(* IEC 61131-3 sources: codesys-framework/txt/application/WeVe Core (library)/30 Module/FB_Module/Properties, 4 files *)

(* ---- Busy.prop.st ---- *)
PROPERTY Busy : BOOL

// --- BEGIN IMPLEMENTATION ---

// ----------- GET -----------
VAR
END_VAR

// -- BEGIN IMPLEMENTATION GET --
Busy := _xBusy;

(* ---- Enabled.prop.st ---- *)
PROPERTY Enabled : BOOL

// --- BEGIN IMPLEMENTATION ---

// ----------- GET -----------
VAR
END_VAR

// -- BEGIN IMPLEMENTATION GET --
Enabled := _xEnabled;

(* ---- Homed.prop.st ---- *)
PROPERTY Homed : BOOL

// --- BEGIN IMPLEMENTATION ---

// ----------- GET -----------
VAR
END_VAR

// -- BEGIN IMPLEMENTATION GET --
Homed := _xHomed;

(* ---- State.prop.st ---- *)
PROPERTY State : E_ModuleStates

// --- BEGIN IMPLEMENTATION ---

// ----------- GET -----------
VAR
END_VAR

// -- BEGIN IMPLEMENTATION GET --
State := _eState;
